// SIMATIC S7-200 project (STEP 7-Micro/WIN), CPU 224XP CN REL 02.01

SYMBOL_TABLE ????1
C_1              VD100
C_0              VD110
x1               VD180
r_k              VD190
u_k              VD150
x2               VD170
x1_1             VD200
N                VD210
K1               VD220
K2               VD230
END_SYMBOL_TABLE

ORGANIZATION_BLOCK ???:OB1
TITLE=????
BEGIN
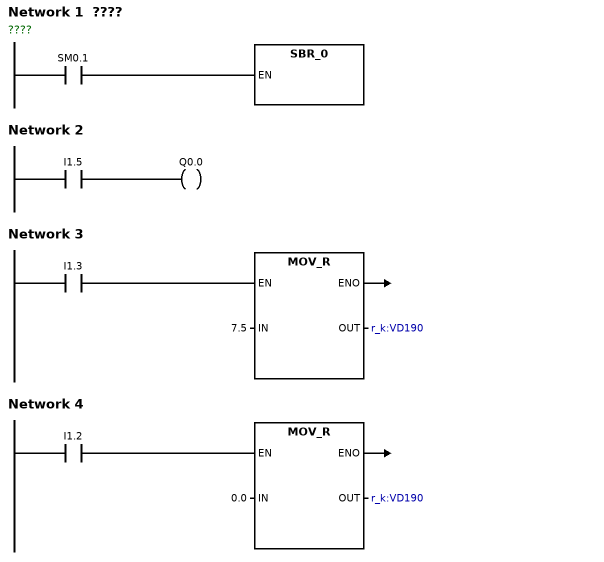
Network 1 // ????
// ????
LD     SM0.1
CALL   SBR_0:SBR0
Network 2
LD     I1.5
=      Q0.0
Network 3
LD     I1.3
MOVR   7.5, r_k:VD190
Network 4
LD     I1.2
MOVR   0.0, r_k:VD190
END_ORGANIZATION_BLOCK

SUBROUTINE_BLOCK SBR_0:SBR0
TITLE=?????
BEGIN
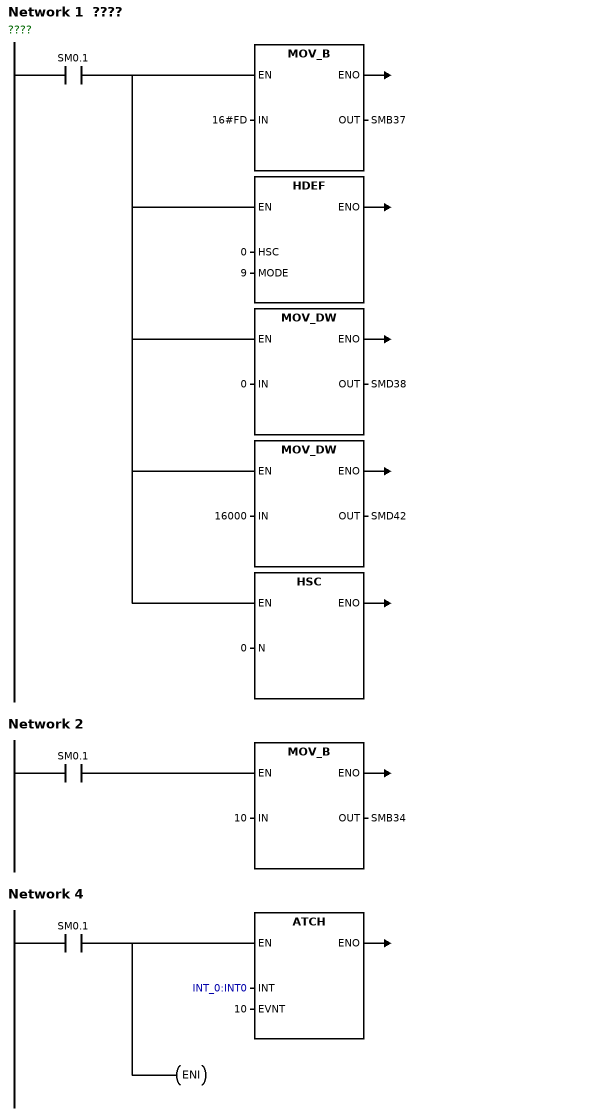
Network 1 // ????
// ????
LD     SM0.1
MOVB   16#FD, SMB37
HDEF   0, 9
MOVD   0, SMD38
MOVD   16000, SMD42
HSC    0
Network 2
LD     SM0.1
MOVB   10, SMB34
Network 4
LD     SM0.1
ATCH   INT_0:INT0, 10
ENI
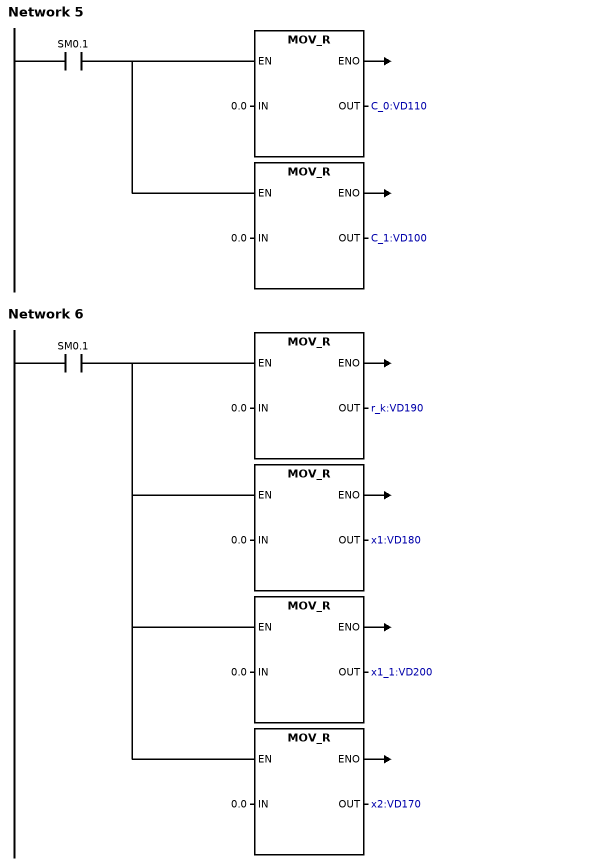
Network 5
LD     SM0.1
MOVR   0.0, C_0:VD110
MOVR   0.0, C_1:VD100
Network 6
LD     SM0.1
MOVR   0.0, r_k:VD190
MOVR   0.0, x1:VD180
MOVR   0.0, x1_1:VD200
MOVR   0.0, x2:VD170
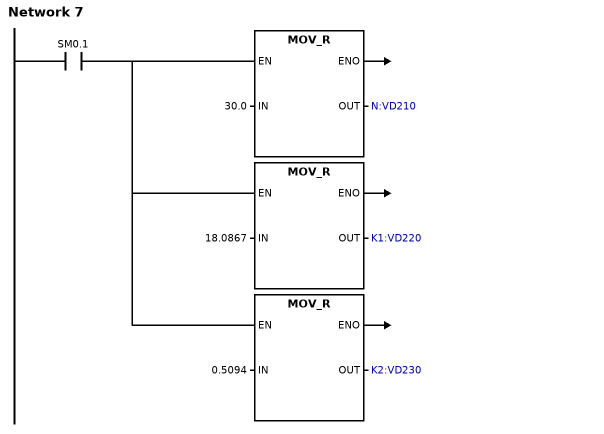
Network 7
LD     SM0.1
MOVR   30.0, N:VD210
MOVR   18.0867, K1:VD220
MOVR   0.5094, K2:VD230
END_SUBROUTINE_BLOCK

INTERRUPT_BLOCK INT_0:INT0
TITLE=??????
BEGIN
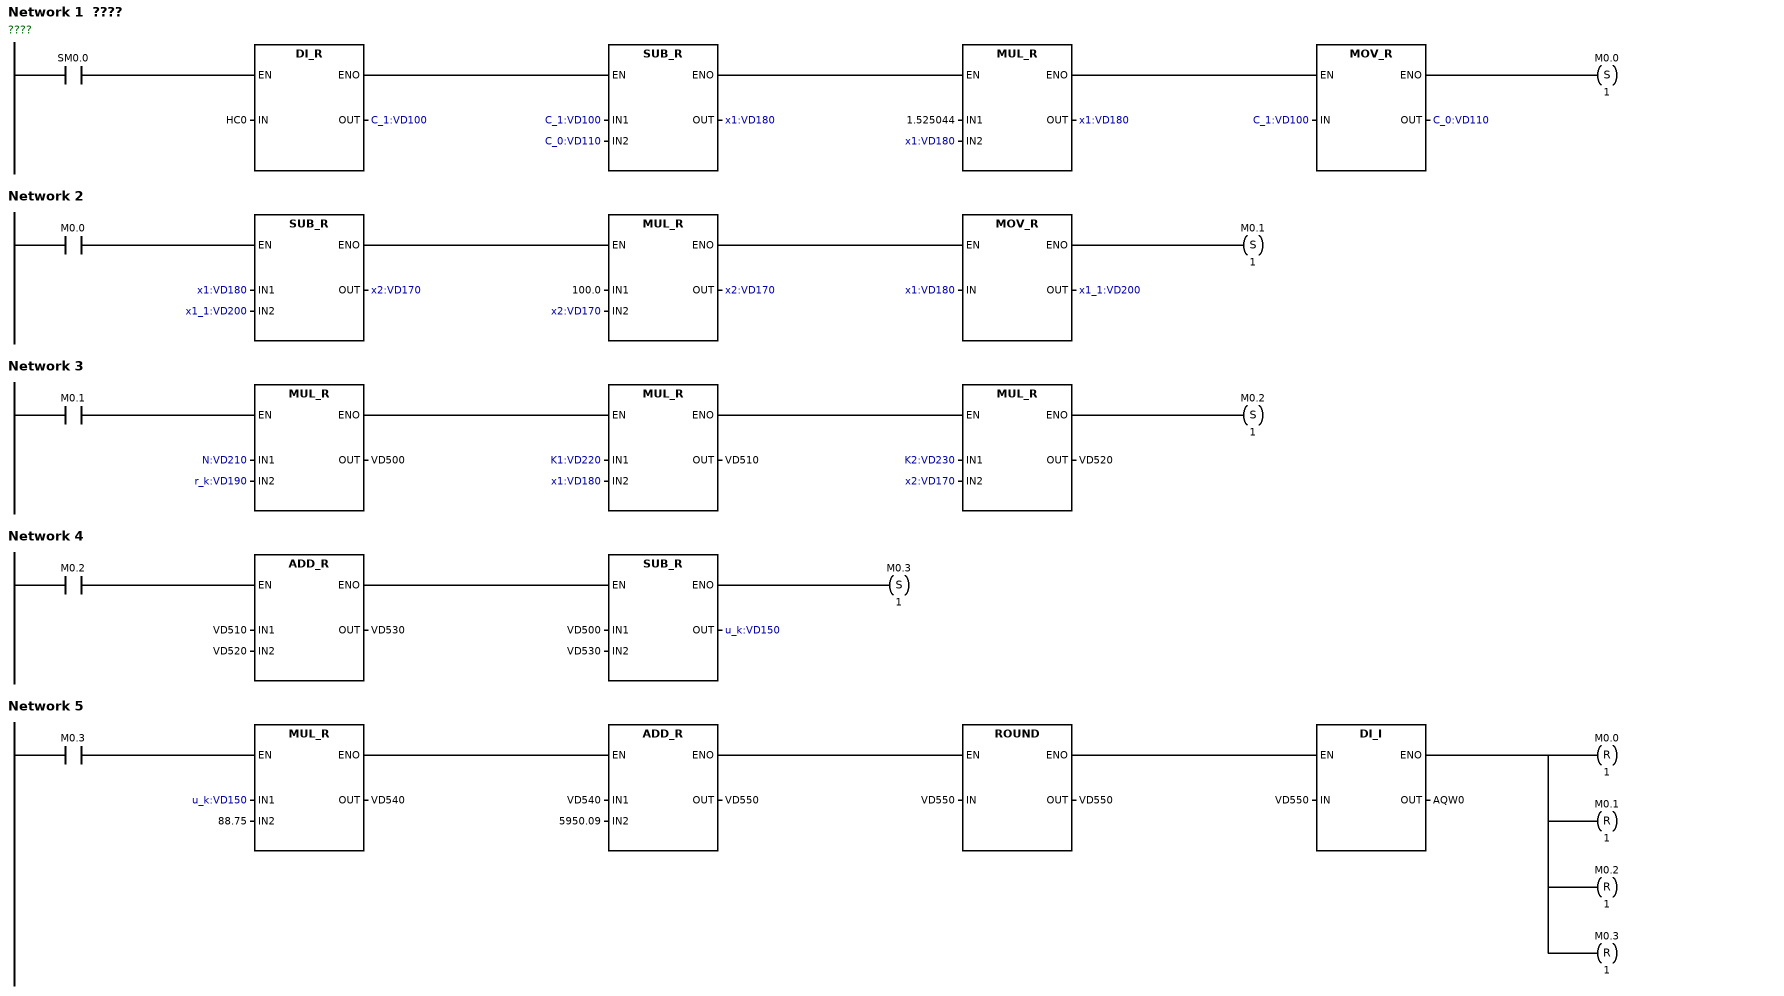
Network 1 // ????
// ????
LD     SM0.0
DTR    HC0, C_1:VD100
AENO
MOVR   C_1:VD100, x1:VD180
AENO
-R     C_0:VD110, x1:VD180
AENO
*R     1.525044, x1:VD180
AENO
MOVR   C_1:VD100, C_0:VD110
AENO
S      M0.0, 1
Network 2
LD     M0.0
MOVR   x1:VD180, x2:VD170
AENO
-R     x1_1:VD200, x2:VD170
AENO
*R     100.0, x2:VD170
AENO
MOVR   x1:VD180, x1_1:VD200
AENO
S      M0.1, 1
Network 3
LD     M0.1
MOVR   N:VD210, VD500
AENO
*R     r_k:VD190, VD500
AENO
MOVR   K1:VD220, VD510
AENO
*R     x1:VD180, VD510
AENO
MOVR   K2:VD230, VD520
AENO
*R     x2:VD170, VD520
AENO
S      M0.2, 1
Network 4
LD     M0.2
MOVR   VD510, VD530
AENO
+R     VD520, VD530
AENO
MOVR   VD500, u_k:VD150
AENO
-R     VD530, u_k:VD150
AENO
S      M0.3, 1
Network 5
LD     M0.3
MOVR   u_k:VD150, VD540
AENO
*R     88.75, VD540
AENO
MOVR   VD540, VD550
AENO
+R     5950.09, VD550
AENO
ROUND  VD550, VD550
AENO
DTI    VD550, AQW0
AENO
R      M0.0, 1
R      M0.1, 1
R      M0.2, 1
R      M0.3, 1
END_INTERRUPT_BLOCK
